SUBAPPLICATION Uebung_149b (* Übung zu ETP empfangen (PGN 0x1EF00, 4000 Byte), Anzeige im Watch *)
  (* Standard: 61499-2; Description: Copyright (c) 2026 Meisterschulen am Ostbahnhof This program and the accompanying materials are made available under the terms of the Eclipse Public License 2.0 which is available at https://www.eclipse.org/legal/epl-2.0/ SPDX-License-Identifier: EPL-2.0 *)
  (* Version 1.0, 2026-11-17, Franz Höpfinger, Meisterschulen am Ostbahnhof, initial API and implementation and/or initial documentation *)
  PACKAGE Uebungen;
  IMPORT Uebungen::const::Uebung_140_149::Etp::LOGIBUS_ADD;
  IMPORT Uebungen::const::Uebung_140_149::Etp::LOGIBUS_FLT;
  IMPORT isobus::pgn::ISOUSERHOME_e::network;
  IMPORT isobus::pgn::ISO_CAN_NODE::NODE1;
  IMPORT isobus::pgn::const::PgnDef::PGN_PDU1_PropA2;
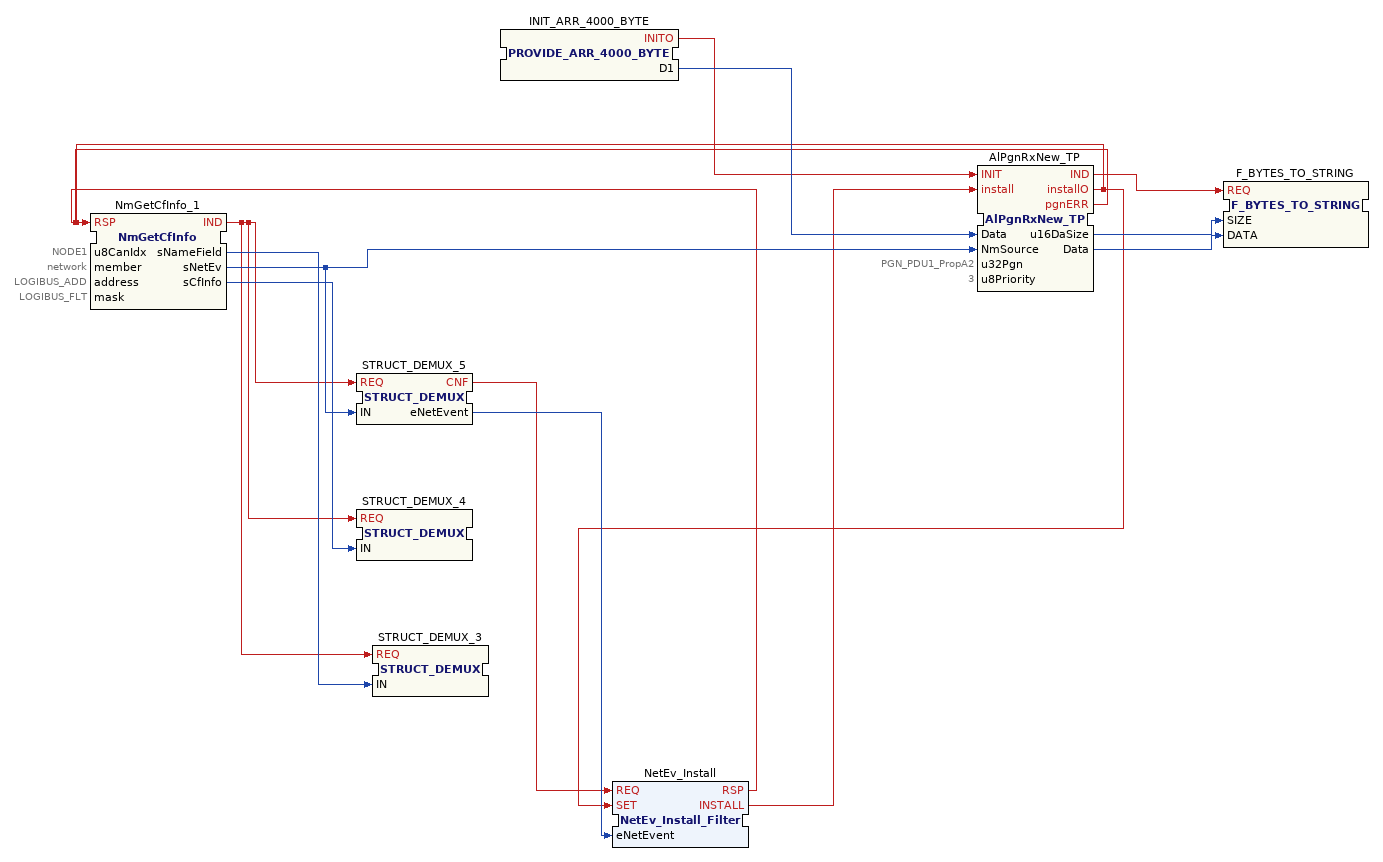
  (* ETP empfangen: PGN PropA2 0x1EF00, 4000 Byte vom anderen logiBUS (Übung 149 oder 149d) Mehr als 1785 Byte gehen per ETP (Extended Transport Protocol), nur an einen Empfänger. Partner: NmGetCfInfo mit network + Filter LOGIBUS_ADD/LOGIBUS_FLT. Puffer 4000 Byte. Watch: u16DaSize = 4000, OVERFLOW = FALSE, Text = ETP-Test 4000 Byte. Firmware ab LOGIBUS 24534469 auf BEIDEN Geräten. *)
  FBS
    STRUCT_DEMUX_3 : eclipse4diac::convert::STRUCT_DEMUX; {SET_ATTRIBUTE(StructuredType, isobus::pgn::NAMEFIELD_T)}
    NmGetCfInfo_1 : isobus::pgn::NmGetCfInfo(u8CanIdx := NODE1, member := network, address := LOGIBUS_ADD, mask := LOGIBUS_FLT);
    STRUCT_DEMUX_4 : eclipse4diac::convert::STRUCT_DEMUX; {SET_ATTRIBUTE(StructuredType, isobus::pgn::CF_INFO_T)}
    STRUCT_DEMUX_5 : eclipse4diac::convert::STRUCT_DEMUX; {SET_ATTRIBUTE(StructuredType, isobus::pgn::ISONETEVENT_T)}
    INIT_ARR_4000_BYTE : eclipse4diac::convert::providers::PROVIDE_ARR_4000_BYTE;
    AlPgnRxNew_TP : isobus::pgn::rx::AlPgnRxNew_TP(u32Pgn := PGN_PDU1_PropA2, u8Priority := 3);
    F_BYTES_TO_STRING : logiBUS::utils::dyn_arr::F_BYTES_TO_STRING;
  END_FBS
  SUBAPPS
    NetEv_Install : MyLib::sys::NetEv_Install_Filter;
  END_SUBAPPS
  EVENT_CONNECTIONS
    NmGetCfInfo_1.IND TO STRUCT_DEMUX_3.REQ;
    NmGetCfInfo_1.IND TO STRUCT_DEMUX_4.REQ;
    NmGetCfInfo_1.IND TO STRUCT_DEMUX_5.REQ;
    INIT_ARR_4000_BYTE.INITO TO AlPgnRxNew_TP.INIT;
    AlPgnRxNew_TP.IND TO F_BYTES_TO_STRING.REQ;
    AlPgnRxNew_TP.installO TO NmGetCfInfo_1.RSP;
    AlPgnRxNew_TP.pgnERR TO NmGetCfInfo_1.RSP;
    STRUCT_DEMUX_5.CNF TO NetEv_Install.REQ;
    NetEv_Install.RSP TO NmGetCfInfo_1.RSP;
    AlPgnRxNew_TP.installO TO NetEv_Install.SET;
    NetEv_Install.INSTALL TO AlPgnRxNew_TP.install;
  END_CONNECTIONS
  DATA_CONNECTIONS
    NmGetCfInfo_1.sNameField TO STRUCT_DEMUX_3.IN;
    NmGetCfInfo_1.sNetEv TO STRUCT_DEMUX_5.IN;
    NmGetCfInfo_1.sCfInfo TO STRUCT_DEMUX_4.IN;
    INIT_ARR_4000_BYTE.D1 TO AlPgnRxNew_TP.Data;
    AlPgnRxNew_TP.u16DaSize TO F_BYTES_TO_STRING.SIZE;
    AlPgnRxNew_TP.Data TO F_BYTES_TO_STRING.DATA;
    STRUCT_DEMUX_5.eNetEvent TO NetEv_Install.eNetEvent;
    NmGetCfInfo_1.sNetEv TO AlPgnRxNew_TP.NmSource;
  END_CONNECTIONS
END_SUBAPPLICATION
